(* CODESYS project P_InstancePath.xml

Project tree, tasks and I/O mapping:
*)

// P_InstancePath
PROPERTY P_InstancePath : STRING
END_PROPERTY
